(* IEC 61131-3 sources: llm-plc-st-eval/data/processed_definitivo/claude-sonnet-4-6/B4/few_shot, 3 files *)

(* ---- ejec_1.st ---- *)
FUNCTION_BLOCK FB_Giro
VAR_INPUT
    btnFwd  : BOOL; (* Boton marcha sentido horario *)
    btnRev  : BOOL; (* Boton marcha sentido antihorario *)
    btnParo : BOOL; (* Boton de paro *)
END_VAR
VAR_OUTPUT
    fwd : BOOL; (* Salida sentido horario *)
    rev : BOOL; (* Salida sentido antihorario *)
END_VAR
VAR
    stateFwd : BOOL; (* Estado interno: motor girando en horario *)
    stateRev : BOOL; (* Estado interno: motor girando en antihorario *)
END_VAR

(* Paro: desactiva ambos sentidos *)
IF btnParo THEN
    stateFwd := FALSE;
    stateRev := FALSE;

(* Arranque horario: solo si el sentido antihorario esta detenido *)
ELSIF btnFwd AND NOT stateRev THEN
    stateFwd := TRUE;

(* Arranque antihorario: solo si el sentido horario esta detenido *)
ELSIF btnRev AND NOT stateFwd THEN
    stateRev := TRUE;
END_IF;

(* Asignacion de salidas; garantia hardware: nunca ambas activas *)
fwd := stateFwd AND NOT stateRev;
rev := stateRev AND NOT stateFwd;

END_FUNCTION_BLOCK

(* ---- ejec_2.st ---- *)
FUNCTION_BLOCK FB_Giro
VAR_INPUT
    btnFwd  : BOOL; (* Boton marcha horaria *)
    btnRev  : BOOL; (* Boton marcha antihoraria *)
    btnParo : BOOL; (* Boton de paro *)
END_VAR
VAR_OUTPUT
    fwd : BOOL; (* Salida giro horario *)
    rev : BOOL; (* Salida giro antihorario *)
END_VAR

(* Logica de enclavamiento con paso obligatorio por paro *)

(* Paro: desactiva ambas salidas *)
IF btnParo THEN
    fwd := FALSE;
    rev := FALSE;

(* Marcha horaria: solo si rev no esta activa (no se permite inversion directa) *)
ELSIF btnFwd AND NOT rev THEN
    fwd := TRUE;

(* Marcha antihoraria: solo si fwd no esta activa (no se permite inversion directa) *)
ELSIF btnRev AND NOT fwd THEN
    rev := TRUE;
END_IF;

(* Seguridad hardware: garantiza exclusion mutua ante cualquier condicion imprevista *)
IF fwd AND rev THEN
    fwd := FALSE;
    rev := FALSE;
END_IF;

END_FUNCTION_BLOCK

(* ---- ejec_3.st ---- *)
FUNCTION_BLOCK FB_Giro
VAR_INPUT
    btnFwd  : BOOL; (* Boton marcha horaria *)
    btnRev  : BOOL; (* Boton marcha antihoraria *)
    btnParo : BOOL; (* Boton de paro *)
END_VAR
VAR_OUTPUT
    fwd : BOOL; (* Salida giro horario *)
    rev : BOOL; (* Salida giro antihorario *)
END_VAR

(* Paro: desactiva ambas salidas *)
IF btnParo THEN
    fwd := FALSE;
    rev := FALSE;

(* Marcha horaria: solo si rev no esta activa (paso previo por paro obligatorio) *)
ELSIF btnFwd AND NOT rev THEN
    fwd := TRUE;

(* Marcha antihoraria: solo si fwd no esta activa (paso previo por paro obligatorio) *)
ELSIF btnRev AND NOT fwd THEN
    rev := TRUE;
END_IF;

(* Enclavamiento de seguridad: nunca ambas salidas activas simultaneamente *)
IF fwd AND rev THEN
    fwd := FALSE;
    rev := FALSE;
END_IF;
END_FUNCTION_BLOCK
